(* IEC 61131-3 sources: trust-platform/examples/ladder, 2 files *)

(* ---- simple-start-stop.st ---- *)
(*
  Auto-generated from ladder source: simple-start-stop.ladder.json
  Source of truth is the visual file unless migrated fully to ST.
*)
(*
  Auto-generated Ladder Diagram companion (schema v2).
  Source of truth remains the .ladder.json file.
  Generated to support .st-first runtime workflows.
*)

FUNCTION_BLOCK FB_simple_start_stop_LADDER
VAR_EXTERNAL
  StartPB : BOOL;
  StopPB : BOOL;
  MotorRun : BOOL;
  AlarmLamp : BOOL;
END_VAR

VAR
  dfg : BOOL := FALSE; (* Ladder local *)
  test : BOOL := FALSE; (* Ladder local *)
END_VAR

(* Network 0: rung_1 *)
MotorRun := StartPB OR dfg OR test;

(* Network 1: rung_2 *)
AlarmLamp := NOT (StopPB);

END_FUNCTION_BLOCK

(* ---- simple-start-stop.visual.runtime.st ---- *)
(*
  Auto-generated runtime entry for simple-start-stop.ladder.json.
  This wrapper is used to run visual editors through the Structured Text debugger path.
*)

PROGRAM PRG_simple_start_stop_VISUAL
fb_simple_start_stop();
END_PROGRAM

CONFIGURATION CFG_simple_start_stop_VISUAL
VAR_GLOBAL
  fb_simple_start_stop : FB_simple_start_stop_LADDER;
  StartPB AT %IX0.0 : BOOL;
  StopPB AT %IX0.1 : BOOL;
  MotorRun AT %QX0.0 : BOOL;
  AlarmLamp AT %QX0.1 : BOOL;
END_VAR
  RESOURCE RES_simple_start_stop_VISUAL ON PLC
    TASK TASK_simple_start_stop_VISUAL(INTERVAL := T#20ms, PRIORITY := 1);
    PROGRAM PLC_PRG_simple_start_stop WITH TASK_simple_start_stop_VISUAL : PRG_simple_start_stop_VISUAL;
  END_RESOURCE
END_CONFIGURATION
